(* LS Electric XG5000 project: TEXTOK *)
(* PLC LSPLC *)

PROGRAM AddedProgram (* task: 스캔 프로그램 *)
END_PROGRAM

PROGRAM NewProgram (* task: 스캔 프로그램 *)
VAR
    GOTO_INIT : BOOL;
    TRANS : BOOL;
END_VAR
(* SFC body not rendered *)
END_PROGRAM

PROGRAM NativeST (* task: 스캔 프로그램 *)
%MX0 := TRUE;
END_PROGRAM

PROGRAM NativeIL (* task: 스캔 프로그램 *)
LD 1
ST %MW0
END_PROGRAM